TYPE "ST_DigitalInputParCfg"
VERSION : 0.1
   STRUCT
      "SchemaVersion" : UInt := 1;
   END_STRUCT;
END_TYPE
